Staubli VAL3: saveTask.pgx

program saveTask()
begin
  db:libSave()
end
